KUKA KRL program: InspectA.src

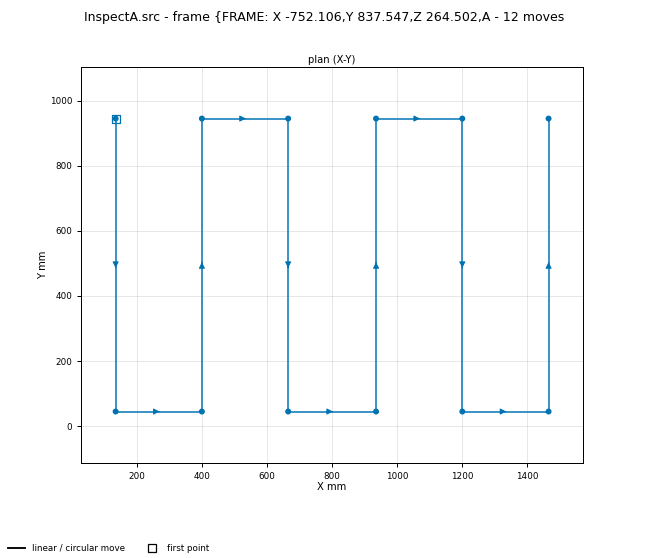
[picture p0: tool path of InspectA.src in frame {FRAME: X -752.106,Y 837.547,Z 264.502,A, 12 of 12 moves have a stored position in this frame; points joined in program order, loops and branches not executed]
&ACCESS RVP
&REL 1
&PARAM TEMPLATE = C:\KRC\Roboter\Template\vorgabe
&PARAM EDITMASK = *
DEF InspectA ( )
EXT BAS (BAS_COMMAND :IN,REAL :IN )


; GLOBAL INTERRUPT DECL 3 WHEN $STOPMESS==TRUE DO IR_STOPM ( )
; INTERRUPT ON 3

;FOLD Initialise and set default speed
BAS (#INITMOV,0)
BAS (#VEL_PTP,100)
BAS (#ACC_PTP,20)
$VEL.CP=0.2
BAS (#TOOL,0)
BAS (#BASE,0)
;ENDFOLD

;;FOLD STARTPOS
;$BWDSTART = FALSE
;PDAT_ACT = PDEFAULT
;BAS(#PTP_DAT)
;FDAT_ACT = {TOOL_NO 0,BASE_NO 0,IPO_FRAME #BASE}
;BAS(#FRAMES)
;;ENDFOLD

$ADVANCE = 5

;FOLD ---- Quickly skip BCO ----
; PTP $AXIS_ACT
;ENDFOLD

;FOLD ---- GO HOME ----
; PTP {A1 0.000, A2 -90.000, A3 90.000, A4 0.000, A5 0.000, A6 0.000, E1 0, E2 0, E3 0, E4 0, E5 0, E6 0}
;ENDFOLD


; Program generated by VerticalBot Studio for KUKA KR 22 R1610 on 25/10/2026 12:00:00
; Using nominal kinematics.
; ---- Setting reference (Base) ----
$BASE = {FRAME: X -752.106,Y 837.547,Z 264.502,A 0.000,B 0.000,C 32.841}
; --------------------------
; ---- Setting tool (TCP) ----
; TOOL_DATA[2] = {FRAME: X 245.414,Y 0.000,Z 424.009,A 0.000,B 36.800,C 0.000}
$TOOL = {FRAME: X 245.414,Y 0.000,Z 424.009,A 0.000,B 36.800,C 0.000}
; $TOOL = TOOL_DATA[2]
; --------------------------
LIN {X 135.000,Y 945.000,Z 9.786,A -90.000,B 0.000,C -180.000}
LIN {X 135.000,Y 45.000,Z 10.000,A -90.000,B 0.000,C -180.000}
LIN {X 400.000,Y 45.000,Z 10.000,A -90.000,B 0.000,C -180.000}
LIN {X 400.000,Y 945.000,Z 10.000,A -90.000,B 0.000,C -180.000}
LIN {X 665.000,Y 945.000,Z 10.000,A -90.000,B 0.000,C -180.000}
LIN {X 665.000,Y 45.000,Z 10.000,A -90.000,B 0.000,C 180.000}
LIN {X 935.000,Y 45.000,Z 10.000,A -90.000,B 0.000,C 180.000}
LIN {X 935.000,Y 945.000,Z 10.000,A -90.000,B 0.000,C 180.000}
LIN {X 1200.000,Y 945.000,Z 10.000,A -90.000,B 0.000,C -180.000}
LIN {X 1200.000,Y 45.000,Z 10.000,A -90.000,B 0.000,C -180.000}
LIN {X 1465.000,Y 45.000,Z 10.000,A -90.000,B 0.000,C 180.000}
LIN {X 1465.000,Y 945.000,Z 10.000,A -90.000,B 0.000,C -180.000}
END
